(* IEC 61131-3 sources: Gen-AI/final/Gen-AI_v1.0_submission/A2_框架源码/agent/logs/full34_fixture/E3_P04_1_42/tools/candidate_1/fixture_compile, 1 file *)

(* ---- source.st ---- *)
FUNCTION_BLOCK FB_P04
VAR_INPUT
    VISCOSITY_OK : BOOL;
    PASTE_E_STOP_NC : BOOL;
    DebounceTime : TIME;
    CycleTime : TIME;
END_VAR
VAR_OUTPUT
    VFD_RUN : BOOL;
    PUMP_MAINT_DUE : BOOL;
    PUMP_RUNTIME_ACC : LTIME;
END_VAR
(* Add a VAR block for internal state/timers before the implementation, if needed. *)
(* SKELETON ONLY: replace this RETURN with scan logic and required initial state. *)
RETURN;
END_FUNCTION_BLOCK

(* FIXTURE_COMPILE_FAIL *)
